Staubli VAL3: main.pgx

program main()
begin
  close(tCurrentTool)
  pPointRx.config.shoulder = lefty
  pPointRx.config.elbow = epositive
  pPointRx.config.wrist = wpositive
  pPointRx2.config.shoulder = lefty
  pPointRx2.config.elbow = epositive
  pPointRx2.config.wrist = wpositive
  mCurrentSpeed.tvel = 100.00
  mCurrentSpeed.blend = joint
  mCurrentSpeed.reach = 0.010
  mCurrentSpeed.leave = 0.010
  // Program FeatureTest start
  // Program generated by VerticalBot Studio for Staubli RX160 on 25/10/2026 12:00:00
  // Using nominal kinematics.
  mCurrentSpeed.tvel = 300.000
  mCurrentSpeed.reach = 5.000
  mCurrentSpeed.leave = 5.000
  call MoveJoint(10.00000,20.00000,90.00000,30.00000,45.00000,60.00000)
  call MoveLine(1077.300,-56.172,837.243,-146.156,25.288,-102.118)
  call MoveCirc(1005.190,-118.362,847.372,-147.806,26.655,-97.799,1002.360,-324.842,854.563,-153.015,33.232,-88.833)
  mCurrentSpeed.tvel = 50.000
  mCurrentSpeed.reach = 0.000
  mCurrentSpeed.leave = 0.000
  call MoveLine(1077.300,-56.172,837.243,-146.156,25.288,-102.118)
  mCurrentSpeed.reach = -1.000
  mCurrentSpeed.leave = -1.000
  mCurrentSpeed.tvel = 300.000
  call MoveLine(1005.190,-118.362,847.372,-147.806,26.655,-97.799)
  Output[3]=true
  DO_GRIP=false
  watch(Input[5]==true)
  watch(DI_PART==true,2000.0)
  delay(0.500)
  // a comment line
  popUpMsg("Hello operator")
  //call prog:MyFunc()
  //call prog:SetRPM(5000)
  RAW_CODE_LINE
  //call prog:SubPick()
  // Attach to Tool 1
  call MoveJoint(10.00000,20.00000,90.00000,30.00000,45.00000,60.00000)
  popUpMsg("Paused. Press OK to continue")

  waitEndMove()
  // Program FeatureTest end

end
